Universal Robots PolyScope program: step5d_autotuner_xy_no_contact_diagnostic_v1.urp

Program step5d_autotuner_xy_no_contact_diagnostic_v1 (installation=default directory=/programs/andyl/kunwei/step5 createdIn=5.11.9.1010452 lastSavedIn=5.11.9.1010452 robotSerialNumber=20225200364)
Calibrated DH parameters: a=[0.00002, -0.569483, -0.54992, -0.00001, -0.000036, 0]; d=[0.180894, -146.691669, 192.918669, -46.053088, 0.119778, 0.115602]; alpha=[1.571425, -0.001534, 0.003359, 1.568739, -1.571477, 0]; deltaTheta=[0, 0.376258, -0.101074, -0.275185, -0.000002, 0]
Robot Program (runOnlyOnce=true)
  Script file /programs/andyl/kunwei/step5/step5d_autotuner_xy_no_contact_diagnostic_v1.script
    | # VERSION: 20260815_STEP5D_AUTOTUNER_XY_NO_CONTACT_DIAGNOSTIC_V1
    | # PURPOSE: one-shot 60 s autotuner absolute-XY, startup fixed-Z/orientation, no contact/search/force control.
    | # WIRE: input float 24 force norm, 25 torque norm, 26 heartbeat, 27 sensor fresh, 28 abort, 29 phase, 37..42 qdot, 43 valid, 44 path time, 47 layout=725.
    | # LIFECYCLE: guarded preposition -> one PATH -> guarded path-origin -> startup Home -> stationary. Faults zero/abort without recovery motion.
    | 
    | def codex_abs(x):
    |   if x < 0:
    |     return -x
    |   end
    |   return x
    | end
    | 
    | def codex_guard_reason(last_heartbeat, stale_s):
    |   local heartbeat = read_input_float_register(26)
    |   local sensor_ok = read_input_float_register(27)
    |   local abort_reason = read_input_float_register(28)
    |   local force_norm = read_input_float_register(24)
    |   local torque_norm = read_input_float_register(25)
    |   if sensor_ok < 0.5:
    |     return [2.0, heartbeat, stale_s]
    |   elif abort_reason > 0.5:
    |     return [abort_reason, heartbeat, stale_s]
    |   elif force_norm > 6.0:
    |     return [6.0, heartbeat, stale_s]
    |   elif torque_norm > 0.5:
    |     return [7.0, heartbeat, stale_s]
    |   end
    |   if heartbeat == last_heartbeat:
    |     stale_s = stale_s + get_steptime()
    |   else:
    |     stale_s = 0.0
    |   end
    |   if stale_s > 1.0:
    |     return [2.0, heartbeat, stale_s]
    |   end
    |   return [0.0, heartbeat, stale_s]
    | end
    | 
    | def codex_guarded_xy_move(target_pose, stage_code, last_heartbeat, stale_s):
    |   write_output_float_register(35, stage_code)
    |   local reason = 0.0
    |   local elapsed = 0.0
    |   while reason == 0.0 and elapsed < 75.0:
    |     local guard = codex_guard_reason(last_heartbeat, stale_s)
    |     reason = guard[0]
    |     last_heartbeat = guard[1]
    |     stale_s = guard[2]
    |     local current = get_actual_tcp_pose()
    |     local ex = target_pose[0] - current[0]
    |     local ey = target_pose[1] - current[1]
    |     local distance = sqrt(ex*ex + ey*ey)
    |     write_output_float_register(36, distance)
    |     if reason == 0.0:
    |       if distance <= 0.00020:
    |         stopl(0.1)
    |         return [0.0, last_heartbeat, stale_s]
    |       end
    |       local speed = 2.0*distance
    |       if speed > 0.003:
    |         speed = 0.003
    |       end
    |       local vx = speed*ex/distance
    |       local vy = speed*ey/distance
    |       speedl([vx, vy, 0.0, 0.0, 0.0, 0.0], 0.05, 0.002)
    |     end
    |     elapsed = elapsed + get_steptime()
    |   end
    |   stopl(0.1)
    |   if reason == 0.0:
    |     reason = 15.0
    |   end
    |   return [reason, last_heartbeat, stale_s]
    | end
    | 
    | def codex_step5d_autotuner_xy_no_contact_diagnostic_v1():
    |   write_output_float_register(28, 0.0)
    |   write_output_float_register(35, 20.0)
    |   write_output_float_register(47, 0.0)
    |   local reason = 0.0
    |   local last_heartbeat = read_input_float_register(26)
    |   local stale_s = 0.0
    |   local wait_s = 0.0
    |   local fresh_count = 0.0
    |   while reason == 0.0 and fresh_count < 2.0 and wait_s < 30.0:
    |     local guard0 = codex_guard_reason(last_heartbeat, stale_s)
    |     reason = guard0[0]
    |     if guard0[1] != last_heartbeat and read_input_float_register(27) >= 0.5:
    |       fresh_count = fresh_count + 1.0
    |     end
    |     last_heartbeat = guard0[1]
    |     stale_s = guard0[2]
    |     wait_s = wait_s + get_steptime()
    |     sync()
    |   end
    |   if reason == 0.0 and fresh_count < 2.0:
    |     reason = 2.0
    |   end
    | 
    |   local session_home = get_actual_tcp_pose()
    |   local path_origin = p[0.487795411149049, 0.129326792700607, session_home[2], session_home[3], session_home[4], session_home[5]]
    |   if reason == 0.0:
    |     local moved0 = codex_guarded_xy_move(path_origin, 30.0, last_heartbeat, stale_s)
    |     reason = moved0[0]
    |     last_heartbeat = moved0[1]
    |     stale_s = moved0[2]
    |   end
    | 
    |   if reason == 0.0:
    |     write_output_float_register(35, 25.0)
    |     local path_s = 0.0
    |     local accepted = False
    |     while reason == 0.0 and read_input_float_register(29) < 1.5 and path_s < 65.0:
    |       local guard1 = codex_guard_reason(last_heartbeat, stale_s)
    |       reason = guard1[0]
    |       last_heartbeat = guard1[1]
    |       stale_s = guard1[2]
    |       local valid = read_input_float_register(43)
    |       local layout = read_input_float_register(47)
    |       local q0 = read_input_float_register(37)
    |       local q1 = read_input_float_register(38)
    |       local q2 = read_input_float_register(39)
    |       local q3 = read_input_float_register(40)
    |       local q4 = read_input_float_register(41)
    |       local q5 = read_input_float_register(42)
    |       write_output_float_register(36, q0)
    |       write_output_float_register(37, q1)
    |       write_output_float_register(38, q2)
    |       write_output_float_register(39, q3)
    |       write_output_float_register(40, q4)
    |       write_output_float_register(41, q5)
    |       write_output_float_register(42, valid)
    |       write_output_float_register(43, read_input_float_register(44))
    |       write_output_float_register(46, layout)
    |       if reason == 0.0:
    |         if valid >= 0.5 and codex_abs(layout-725.000) < 0.001 and codex_abs(q0) <= 0.15 and codex_abs(q1) <= 0.15 and codex_abs(q2) <= 0.15 and codex_abs(q3) <= 0.15 and codex_abs(q4) <= 0.15 and codex_abs(q5) <= 0.15:
    |           accepted = True
    |           write_output_float_register(47, 1.0)
    |           speedj([q0,q1,q2,q3,q4,q5], 0.05, 0.002)
    |         elif path_s < 1.0 and not accepted:
    |           sync()
    |         else:
    |           reason = 12.0
    |         end
    |       end
    |       path_s = path_s + get_steptime()
    |     end
    |     stopj(0.3)
    |     stopl(0.1)
    |     if reason == 0.0 and read_input_float_register(29) < 1.5:
    |       reason = 16.0
    |     end
    |   end
    | 
    |   if reason == 0.0:
    |     local moved1 = codex_guarded_xy_move(path_origin, 40.0, last_heartbeat, stale_s)
    |     reason = moved1[0]
    |     last_heartbeat = moved1[1]
    |     stale_s = moved1[2]
    |   end
    |   if reason == 0.0:
    |     local moved2 = codex_guarded_xy_move(session_home, 41.0, last_heartbeat, stale_s)
    |     reason = moved2[0]
    |   end
    |   stopj(0.3)
    |   stopl(0.1)
    |   write_output_float_register(28, reason)
    |   if reason == 0.0:
    |     sleep(0.5)
    |     write_output_float_register(35, 78.0)
    |   else:
    |     write_output_float_register(35, 90.0)
    |   end
    | end
    | 
    | codex_step5d_autotuner_xy_no_contact_diagnostic_v1()
